(* IEC 61131-3 sources: codesys-api/examples/mqtt_large_payload/st/bcnf_comms, 3 files *)

(* ---- BenchFirstPublish.st ---- *)
FUNCTION_BLOCK BenchFirstPublish
// BCNF's FirstPublish (PLC_BCNF_4_16_26) verbatim, on BcnfComms.MQTT_PUBLISH; topic raw_data -> raw_data_demo/bcnf/raw;
// SysTimeRtcHighResGet -> NowUs() (the demo has no SysTimeRtc reference; the value is not published).
VAR_INPUT
    InterlockData1: STRING(255);
    InterlockData2: STRING(255);
    InterlockData3: STRING(255);
    InterlockData4: STRING(255);
    InterlockData5: STRING(255);
    InterlockData6: STRING(255);
    InterlockData7: STRING(255);
END_VAR
VAR_OUTPUT
    PublishDone: BOOL;                          // Indicates when publish operation completes
END_VAR
VAR
    // ===== MQTT PUBLISHER CORE =====
    publisher1: MQTT.MQTTPublish;
    publisher2: MQTT.MQTTPublish;
    publisher3: MQTT.MQTTPublish;
    publisher4: MQTT.MQTTPublish;
    publisher5: MQTT.MQTTPublish;
    publisher6: MQTT.MQTTPublish;
    publisher7: MQTT.MQTTPublish;

    init: BOOL;                                // One-time initialization flag

    // ===== MESSAGE CONTENT =====
    fullPayload1: STRING(255);
    fullPayload2: STRING(255);
    fullPayload3: STRING(255);
    fullPayload4: STRING(255);
    fullPayload5: STRING(255);
    fullPayload6: STRING(255);
    fullPayload7: STRING(255);

    // ===== PUBLISHING CONTROL =====
    sendTimer: TON;                            // Timer controlling publish frequency
    readyToSend: BOOL;                         // Flag indicating ready to publish

    // ===== MESSAGE STATISTICS =====
    TicCount: UDINT;
    TicCountOld: UDINT;
    TicsPerSecond: REAL;
    totalMessages: UDINT;
    PulseCount: UDINT;
    previousTotalMessages: UDINT;
    messagesPerSecond: REAL;

    // ===== TIMING AND STATE TRACKING =====
    publisher_done_prev: BOOL;
    rateTimer: TON;

    // ===== TIMESTAMP GENERATION =====
    dtNowString: STRING;
    RTC: ULINT;

    Pulse: BOOL;
END_VAR
// ---- implementation ----
// ===== EXPOSE PUBLISH STATE =====
TicCount := TicCount + 1;
PublishDone := publisher1.done;

// ===== ONE-TIME INITIALIZATION =====
IF NOT init THEN
    init := TRUE;
    publisher1.SetMqttInOut(MQTT_IN_OUT := BcnfComms.MQTT_PUBLISH);
    publisher2.SetMqttInOut(MQTT_IN_OUT := BcnfComms.MQTT_PUBLISH);
    publisher3.SetMqttInOut(MQTT_IN_OUT := BcnfComms.MQTT_PUBLISH);
    publisher4.SetMqttInOut(MQTT_IN_OUT := BcnfComms.MQTT_PUBLISH);
    publisher5.SetMqttInOut(MQTT_IN_OUT := BcnfComms.MQTT_PUBLISH);
    publisher6.SetMqttInOut(MQTT_IN_OUT := BcnfComms.MQTT_PUBLISH);
    publisher7.SetMqttInOut(MQTT_IN_OUT := BcnfComms.MQTT_PUBLISH);
END_IF

// ===== PUBLISH TIMING CONTROL =====
sendTimer(IN := NOT sendTimer.Q, PT := T#1000MS);

// ===== MESSAGE PREPARATION =====
IF sendTimer.Q AND NOT readyToSend THEN
    readyToSend := TRUE;
    PulseCount := PulseCount + 1;
    IF Pulse = TRUE THEN
        Pulse := FALSE;
    ELSE
        Pulse := TRUE;
    END_IF
    RTC := NowUs();
    dtNowString := TO_STRING(RTC);

    fullPayload1 := InterlockData1;
    fullPayload2 := InterlockData2;
    fullPayload3 := InterlockData3;
    fullPayload4 := InterlockData4;
    fullPayload5 := InterlockData5;
    fullPayload6 := InterlockData6;
    fullPayload7 := InterlockData7;

    IF LEN(fullPayload1) = 0 THEN
        readyToSend := FALSE;
    END_IF;
END_IF;

// ===== PUBLISH COMPLETION TRACKING =====
IF (publisher1.done OR LEN(fullPayload1) = 0) AND
   (publisher2.done OR LEN(fullPayload2) = 0) AND
   (publisher3.done OR LEN(fullPayload3) = 0) AND
   (publisher4.done OR LEN(fullPayload4) = 0) AND
   (publisher5.done OR LEN(fullPayload5) = 0) AND
   (publisher6.done OR LEN(fullPayload6) = 0) AND
   (publisher7.done OR LEN(fullPayload7) = 0) THEN
    IF NOT publisher_done_prev THEN
        totalMessages := totalMessages + 1;
    END_IF;
    PublishDone := TRUE;
ELSE
    PublishDone := FALSE;
END_IF;

publisher_done_prev := PublishDone;

// ===== PUBLISH STATE RESET =====
IF PublishDone THEN
    readyToSend := FALSE;
END_IF;

// ===== PUBLISHING RATE MONITORING =====
rateTimer(IN := NOT rateTimer.Q, PT := T#500MS);
IF rateTimer.Q THEN
    messagesPerSecond := TO_REAL(totalMessages - previousTotalMessages) / 2.0;
    previousTotalMessages := totalMessages;
    TicsPerSecond := TO_REAL(TicCount - TicCountOld) / 2.0;
    TicCountOld := TicCount;
END_IF;

// ===== MQTT PUBLISH OPERATION =====
publisher1(
    Topic := ADR('raw_data_demo/bcnf/raw'),
    PayloadString := ADR(fullPayload1),
    PublishAsString := TRUE,
    QoSin := MQTT.QoS.AtMostOnce,
    MRetain := FALSE,
    send := readyToSend AND (LEN(fullPayload1) > 0));

publisher2(
    Topic := ADR('raw_data_demo/bcnf/raw'),
    PayloadString := ADR(fullPayload2),
    PublishAsString := TRUE,
    QoSin := MQTT.QoS.AtMostOnce,
    MRetain := FALSE,
    send := readyToSend AND (LEN(fullPayload2) > 0));

publisher3(
    Topic := ADR('raw_data_demo/bcnf/raw'),
    PayloadString := ADR(fullPayload3),
    PublishAsString := TRUE,
    QoSin := MQTT.QoS.AtMostOnce,
    MRetain := FALSE,
    send := readyToSend AND (LEN(fullPayload3) > 0));

publisher4(
    Topic := ADR('raw_data_demo/bcnf/raw'),
    PayloadString := ADR(fullPayload4),
    PublishAsString := TRUE,
    QoSin := MQTT.QoS.AtMostOnce,
    MRetain := FALSE,
    send := readyToSend AND (LEN(fullPayload4) > 0));

publisher5(
    Topic := ADR('raw_data_demo/bcnf/raw'),
    PayloadString := ADR(fullPayload5),
    PublishAsString := TRUE,
    QoSin := MQTT.QoS.AtMostOnce,
    MRetain := FALSE,
    send := readyToSend AND (LEN(fullPayload5) > 0));

publisher6(
    Topic := ADR('raw_data_demo/bcnf/raw'),
    PayloadString := ADR(fullPayload6),
    PublishAsString := TRUE,
    QoSin := MQTT.QoS.AtMostOnce,
    MRetain := FALSE,
    send := readyToSend AND (LEN(fullPayload6) > 0));

publisher7(
    Topic := ADR('raw_data_demo/bcnf/raw'),
    PayloadString := ADR(fullPayload7),
    PublishAsString := TRUE,
    QoSin := MQTT.QoS.AtMostOnce,
    MRetain := FALSE,
    send := readyToSend AND (LEN(fullPayload7) > 0));

// ------------------------- //
// ------------------------- //
// ------------------------- //
// ------------------------- //
// ------------------------- //

(* ---- BenchFirstSubscription.st ---- *)
FUNCTION_BLOCK BenchFirstSubscription
// BCNF's FirstSubscription (PLC_BCNF_4_16_26) verbatim, on BcnfComms.MQTT_SUBSCRIBE and bench topics:
// plc_commands/CONC-BCNF-PLC -> raw_data_demo/bcnf/commands, plc_status/CONC -> raw_data_demo/bcnf/status.
VAR_INPUT
END_VAR
VAR_OUTPUT
END_VAR
VAR
	// ===== MQTT SUBSCRIPTION COMPONENTS =====
	collector: MQTT.CallbackCollector;          // Manages multiple callback receivers
	SUB1: MQTT.MQTTSubscribe;                   // Main MQTT subscription function block
	receiver: MQTT.ReceiveString;               // String message receiver/parser

	// ===== READY STATE SUBSCRIPTION =====
	collectorReady: MQTT.CallbackCollector;     // Callback collector for ready messages
	SUB2: MQTT.MQTTSubscribe;                   // Ready state subscription function block
	receiverReady: MQTT.ReceiveString;          // Ready state message receiver/parser

	// ===== INITIALIZATION =====
	init: BOOL;
END_VAR
// ---- implementation ----
// ===== ONE-TIME INITIALIZATION =====
IF NOT init THEN
	init := TRUE;

	SUB1.SetMqttInOut(MQTT_IN_OUT := BcnfComms.MQTT_SUBSCRIBE);
	collector.put(instance := receiver);
	receiver.initAsFindTopic(
		compString := ADR('raw_data_demo/bcnf/commands'),
		returnHit := TRUE
	);

	SUB2.SetMqttInOut(MQTT_IN_OUT := BcnfComms.MQTT_SUBSCRIBE);
	collectorReady.put(instance := receiverReady);
	receiverReady.initAsFindTopic(
		compString := ADR('raw_data_demo/bcnf/status'),
		returnHit := TRUE
	);

END_IF;

// ===== ACTIVE SUBSCRIPTION =====
SUB1(
	Subscribe := TRUE,
	Topic := ADR('raw_data_demo/bcnf/commands'),
	QoSSubscribe := MQTT.QoS.ExactlyOnce,
	ExpectingString := TRUE,
	Callback := collector
);

SUB2(
	Subscribe := TRUE,
	Topic := ADR('raw_data_demo/bcnf/status'),
	QoSSubscribe := MQTT.QoS.ExactlyOnce,
	ExpectingString := TRUE,
	Callback := collectorReady
);

(* ---- BcnfComms.st ---- *)
PROGRAM BcnfComms
// BCNF's MQTT path (PLC_BCNF_4_16_26: POU1, FirstSubscription, FirstPublish) on the bench, nearly verbatim: two client
// connections in one PLC (PUB and SUB, both called every scan), CallbackCollector + ReceiveString subscriptions at
// QoS 2, seven QoS 0 string publishers once a second, plus one MQTTState on the PUB connection. Topics are moved under
// raw_data_demo/bcnf/. Idle (both clients disabled) unless IsEnabled; bcnf_test.py drives it.
VAR
	IsEnabled : BOOL;                       // written online
	BrokerUrl : STRING(250) := '192.168.50.240:1883';
	MQTT_PUBLISH : MQTT.MQTT_IN_OUT;
	MQTT_SUBSCRIBE : MQTT.MQTT_IN_OUT;
	FirstSubscription : BenchFirstSubscription;
	FirstPublish : BenchFirstPublish;
	currentMessage : STRING(255);
	CurrentMqttMessageReady : STRING(255);
	// What bcnf_test.py reads
	PubConnected : BOOL;
	SubConnected : BOOL;
	LastMessage : STRING(255);
	LastReady : STRING(255);
	CommandChanges : UDINT;                 // currentMessage changed: one per command when commands are paced
	ReadyChanges : UDINT;
	// The seven interlock strings BCNF publishes, here changing every scan
	Data : ARRAY[1..7] OF STRING(255);
	Scan : UDINT;
	Index : INT;
	// MQTTState (its request now also ends on Rejected)
	StateFlag : BOOL;                       // written online: each change publishes flag:on / flag:off at QoS 1
	StateBlock : MQTT.MQTTState;
	StateTopic : STRING(64) := 'raw_data_demo/bcnf/state';
	StateName : STRING(16) := 'flag';
	StateOn : STRING(8) := 'on';
	StateOff : STRING(8) := 'off';
	IsStateReady : BOOL;
	// Not in BCNF: a '#' subscription, which must also match its parent level (raw_data_demo/bcnf/wild itself)
	WildSub : MQTT.MQTTSubscribe;
	WildCollector : MQTT.CallbackCollector;
	WildReceiver : MQTT.ReceiveString;          // exactly raw_data_demo/bcnf/wild (ReceiveString compares the whole topic)
	WildChildReceiver : MQTT.ReceiveString;     // exactly raw_data_demo/bcnf/wild/child
	LastWildChild : STRING(255);
	IsWildReady : BOOL;
	WildMessage : STRING(255);
	LastWild : STRING(255);
	WildChanges : UDINT;
END_VAR
// ---- implementation ----
// BCNF calls both clients every scan (its subscriptionInitialized flag is never set); so does this, with ENABLE
// following IsEnabled so that disabling disconnects them
MQTT_PUBLISH.ClientID := 'BENCH_BCNF_PUB';
MQTT_PUBLISH.clientFB(MQTT_IN_OUT := MQTT_PUBLISH, ENABLE := IsEnabled, URL := BrokerUrl, TIMEOUT := T#10S, TLS := FALSE);
MQTT_SUBSCRIBE.ClientID := 'BENCH_BCNF_SUB';
MQTT_SUBSCRIBE.clientFB(MQTT_IN_OUT := MQTT_SUBSCRIBE, ENABLE := IsEnabled, URL := BrokerUrl, TIMEOUT := T#10S, TLS := FALSE);
PubConnected := MQTT_PUBLISH.BROKER_CONNECTED;
SubConnected := MQTT_SUBSCRIBE.BROKER_CONNECTED;
IF NOT IsEnabled THEN
	RETURN;
END_IF

FirstSubscription();
currentMessage := FirstSubscription.receiver.MQTTReceived;
CurrentMqttMessageReady := FirstSubscription.receiverReady.MQTTReceived;
IF currentMessage <> LastMessage THEN
	LastMessage := currentMessage;
	CommandChanges := CommandChanges + 1;
END_IF
IF CurrentMqttMessageReady <> LastReady THEN
	LastReady := CurrentMqttMessageReady;
	ReadyChanges := ReadyChanges + 1;
END_IF

Scan := Scan + 1;
FOR Index := 1 TO 7 DO
	Data[Index] := CONCAT(CONCAT('group', INT_TO_STRING(Index)), CONCAT(':', UDINT_TO_STRING(Scan)));
END_FOR
FirstPublish(InterlockData1 := Data[1], InterlockData2 := Data[2], InterlockData3 := Data[3], InterlockData4 := Data[4],
	InterlockData5 := Data[5], InterlockData6 := Data[6], InterlockData7 := Data[7]);

IF NOT IsStateReady THEN
	IsStateReady := TRUE;
	StateBlock.Init(State := ADR(StateFlag), Topic := ADR(StateTopic), StateName := ADR(StateName),
		MQTT_IN_OUT := MQTT_PUBLISH, StateValueOn := ADR(StateOn), StateValueOff := ADR(StateOff),
		QoS := MQTT.QoS.AtLeastOnce, RetainMqtt := FALSE);
END_IF
StateBlock();

IF NOT IsWildReady THEN
	IsWildReady := TRUE;
	WildSub.SetMqttInOut(MQTT_IN_OUT := MQTT_SUBSCRIBE);
	WildCollector.put(instance := WildReceiver);
	WildReceiver.initAsFindTopic(compString := ADR('raw_data_demo/bcnf/wild'), returnHit := TRUE);
	WildCollector.put(instance := WildChildReceiver);
	WildChildReceiver.initAsFindTopic(compString := ADR('raw_data_demo/bcnf/wild/child'), returnHit := TRUE);
END_IF
WildSub(Subscribe := TRUE, Topic := ADR('raw_data_demo/bcnf/wild/#'), QoSSubscribe := MQTT.QoS.AtLeastOnce,
	ExpectingString := TRUE, Callback := WildCollector);
WildMessage := WildReceiver.MQTTReceived;
LastWildChild := WildChildReceiver.MQTTReceived;
IF WildMessage <> LastWild THEN
	LastWild := WildMessage;
	WildChanges := WildChanges + 1;
END_IF
